Fanuc KAREL source: KT00730.KL

PROGRAM KT00730
%NOLOCKGROUP
VAR
  ARG: ARRAY[4] OF INTEGER
  OUT: BOOLEAN
BEGIN
  OUT = UNINIT(ARG)
END KT00730
